Staubli VAL3: do_switch.pgx

public program do_switch(string x_sKey, num x_nIndex)
  local string l_sValue
  local num l_nIOindex
  local bool l_bErr
  local num l_nValue
  local bool l_bResult
begin
  waitEndMove()
  rs:bInSwitch=true
  l_sValue=progTemp:pProgItem[x_sKey].pProgTemplate[x_nIndex].sSwitchItem.sIOValue
  toNum(l_sValue,l_nIOindex,l_bResult)
  call io:getAnaIO(io:aInItem[l_nIOindex].aAio,l_nValue,l_bErr)
  rs:nSetSwitchValue=l_nValue
end
